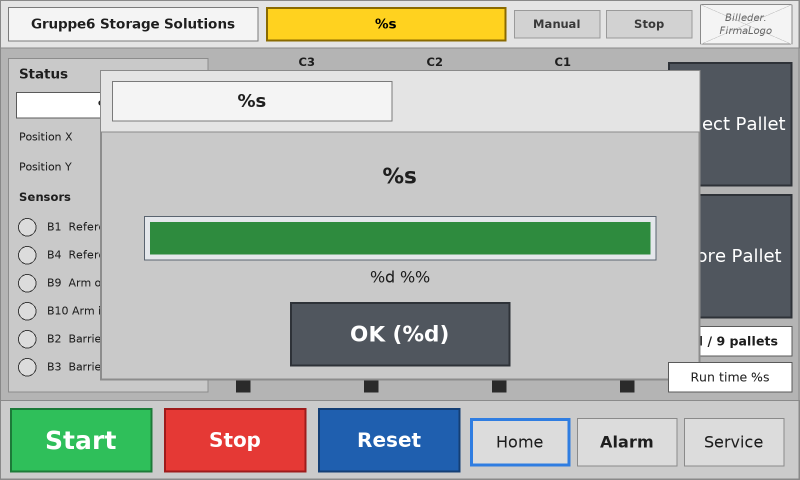
VISUALIZATION Start  // 800x480
    Rectangle (0,0 800x480)
    Rectangle (0,0 800x48)
    Rectangle (8,7 250x34), "Gruppe6 Storage Solutions"
    Rectangle (266,7 150x34), "OP031 Warehouse"
    Rectangle (514,10 86x28), "Manual", colour toggle: MAIN.isManualMode
    Rectangle (606,10 86x28), "Stop", colour toggle: MAIN.isStop
    Rectangle (0,400 800x80)
    RoundedRectangle (10,408 142x64), "Start"
        OnMouseUp: execute { MAIN.isStop := FALSE; }
    RoundedRectangle (164,408 142x64), "Stop"
        OnMouseUp: execute { MAIN.isStop := TRUE; }
    RoundedRectangle (318,408 142x64), "Reset"
        OnMouseUp: execute {
            MAIN.resetRequest := TRUE;   // everything back to Step_10, then homing
        }
    Rectangle (470,418 100x48), "Home"
        OnMouseUp: change screen: Start
    Rectangle (684,418 100x48), "Service"
        OnMouseUp: change screen: Service
    Rectangle (8,58 200x334)
    Rectangle (16,62 184x24), "Status"
    Rectangle (16,124 84x26), "Position X"
    Rectangle (100,124 100x26), "%d", text variable: MAIN.currentPosX
    Rectangle (16,154 84x26), "Position Y"
    Rectangle (100,154 100x26), "%d", text variable: MAIN.currentPosY
    Rectangle (16,186 184x22), "Sensors"
    Ellipse (18,218 18x18), colour toggle: MAIN.B1
    Rectangle (44,214 160x26), "B1 Reference X"
    Ellipse (18,246 18x18), colour toggle: MAIN.B4
    Rectangle (44,242 160x26), "B4 Reference Y (top)"
    Ellipse (18,274 18x18), colour toggle: MAIN.B9
    Rectangle (44,270 160x26), "B9 Arm out"
    Ellipse (18,302 18x18), colour toggle: MAIN.B10
    Rectangle (44,298 160x26), "B10 Arm in"
    Ellipse (18,330 18x18), colour toggle: MAIN.B2
    Rectangle (44,326 160x26), "B2 Barrier in (free)"
    Ellipse (18,358 18x18), colour toggle: MAIN.B3
    Rectangle (44,354 160x26), "B3 Barrier out (free)"
    Rectangle (236,74 14x318)
    Rectangle (364,74 14x318)
    Rectangle (492,74 14x318)
    Rectangle (620,74 14x318)
    Rectangle (236,150 398x10)
    Rectangle (640,120 24x24), "R3"
    Rectangle (236,250 398x10)
    Rectangle (640,220 24x24), "R2"
    Rectangle (236,350 398x10)
    Rectangle (640,320 24x24), "R1"
    Rectangle (277,52 60x20), "C3"
    Rectangle (405,52 60x20), "C2"
    Rectangle (533,52 60x20), "C1"
    Rectangle (265,110 84x40), colour toggle: MAIN.slotOccupied[3,3]
    Rectangle (272,101 70x9), colour toggle: MAIN.slotOccupied[3,3]
    Rectangle (393,110 84x40), colour toggle: MAIN.slotOccupied[2,3]
    Rectangle (400,101 70x9), colour toggle: MAIN.slotOccupied[2,3]
    Rectangle (521,110 84x40), colour toggle: MAIN.slotOccupied[1,3]
    Rectangle (528,101 70x9), colour toggle: MAIN.slotOccupied[1,3]
    Rectangle (265,210 84x40), colour toggle: MAIN.slotOccupied[3,2]
    Rectangle (272,201 70x9), colour toggle: MAIN.slotOccupied[3,2]
    Rectangle (393,210 84x40), colour toggle: MAIN.slotOccupied[2,2]
    Rectangle (400,201 70x9), colour toggle: MAIN.slotOccupied[2,2]
    Rectangle (521,210 84x40), colour toggle: MAIN.slotOccupied[1,2]
    Rectangle (528,201 70x9), colour toggle: MAIN.slotOccupied[1,2]
    Rectangle (265,310 84x40), colour toggle: MAIN.slotOccupied[3,1]
    Rectangle (272,301 70x9), colour toggle: MAIN.slotOccupied[3,1]
    Rectangle (393,310 84x40), colour toggle: MAIN.slotOccupied[2,1]
    Rectangle (400,301 70x9), colour toggle: MAIN.slotOccupied[2,1]
    Rectangle (521,310 84x40), colour toggle: MAIN.slotOccupied[1,1]
    Rectangle (528,301 70x9), colour toggle: MAIN.slotOccupied[1,1]
    RoundedRectangle (668,62 124x124), "Select Pallet"
        OnMouseUp: execute {
            MAIN.awaitingUserInput := TRUE;   // tell the SFC (Step_10): the operator wants to retrieve a pallet
        }
        OnMouseUp: OpenDialog Dialog=SelectPalletDialog, OpenModal=True, OpenCentered=True
    RoundedRectangle (668,194 124x124), "Store Pallet", colour toggle: MAIN.isStorageFull
        OnMouseUp: execute {
            MAIN.storeRequest := TRUE;   // run the pallet in on the conveyor (to B2) and store it in the rack
        }
    Image (700,4 92x40), image: Billeder.FirmaLogo
    Rectangle (16,92 184x26), "%s", text variable: MAIN.statusText
    Rectangle (668,326 124x30), "%d / 9 pallets", text variable: MAIN.palletCount
    Rectangle (100,70 600x310), invisible if: MAIN.hideStorageFull, input disabled if: MAIN.hideStorageFull
    Rectangle (100,70 600x62), invisible if: MAIN.hideStorageFull, input disabled if: MAIN.hideStorageFull
    Rectangle (112,81 200x40), "Warning", invisible if: MAIN.hideStorageFull, input disabled if: MAIN.hideStorageFull
    Rectangle (528,84 160x34), "Storage full", invisible if: MAIN.hideStorageFull, input disabled if: MAIN.hideStorageFull
    Rectangle (120,180 560x60), "Storage is full, remove pallets first", invisible if: MAIN.hideStorageFull, input disabled if: MAIN.hideStorageFull
    RoundedRectangle (290,288 220x64), "OK", invisible if: MAIN.hideStorageFull, input disabled if: MAIN.hideStorageFull
        OnMouseUp: execute {
            MAIN.showStorageFull := FALSE;   // close the message
        }
    Rectangle (100,70 600x310), invisible if: MAIN.hideProgress, input disabled if: MAIN.hideProgress
    Rectangle (100,70 600x62), invisible if: MAIN.hideProgress, input disabled if: MAIN.hideProgress
    Rectangle (112,81 280x40), "%s", text variable: MAIN.progressTitle, invisible if: MAIN.hideProgress, input disabled if: MAIN.hideProgress
    Rectangle (120,148 560x56), "%s", text variable: MAIN.progressText, invisible if: MAIN.hideProgress, input disabled if: MAIN.hideProgress
    Rectangle (144,216 512x44), invisible if: MAIN.hideProgress, input disabled if: MAIN.hideProgress
    Rectangle (150,222 25x32), invisible if: MAIN.progressHide[1], input disabled if: MAIN.progressHide[1]
    Rectangle (175,222 25x32), invisible if: MAIN.progressHide[2], input disabled if: MAIN.progressHide[2]
    Rectangle (200,222 25x32), invisible if: MAIN.progressHide[3], input disabled if: MAIN.progressHide[3]
    Rectangle (225,222 25x32), invisible if: MAIN.progressHide[4], input disabled if: MAIN.progressHide[4]
    Rectangle (250,222 25x32), invisible if: MAIN.progressHide[5], input disabled if: MAIN.progressHide[5]
    Rectangle (275,222 25x32), invisible if: MAIN.progressHide[6], input disabled if: MAIN.progressHide[6]
    Rectangle (300,222 25x32), invisible if: MAIN.progressHide[7], input disabled if: MAIN.progressHide[7]
    Rectangle (325,222 25x32), invisible if: MAIN.progressHide[8], input disabled if: MAIN.progressHide[8]
    Rectangle (350,222 25x32), invisible if: MAIN.progressHide[9], input disabled if: MAIN.progressHide[9]
    Rectangle (375,222 25x32), invisible if: MAIN.progressHide[10], input disabled if: MAIN.progressHide[10]
    Rectangle (400,222 25x32), invisible if: MAIN.progressHide[11], input disabled if: MAIN.progressHide[11]
    Rectangle (425,222 25x32), invisible if: MAIN.progressHide[12], input disabled if: MAIN.progressHide[12]
    Rectangle (450,222 25x32), invisible if: MAIN.progressHide[13], input disabled if: MAIN.progressHide[13]
    Rectangle (475,222 25x32), invisible if: MAIN.progressHide[14], input disabled if: MAIN.progressHide[14]
    Rectangle (500,222 25x32), invisible if: MAIN.progressHide[15], input disabled if: MAIN.progressHide[15]
    Rectangle (525,222 25x32), invisible if: MAIN.progressHide[16], input disabled if: MAIN.progressHide[16]
    Rectangle (550,222 25x32), invisible if: MAIN.progressHide[17], input disabled if: MAIN.progressHide[17]
    Rectangle (575,222 25x32), invisible if: MAIN.progressHide[18], input disabled if: MAIN.progressHide[18]
    Rectangle (600,222 25x32), invisible if: MAIN.progressHide[19], input disabled if: MAIN.progressHide[19]
    Rectangle (625,222 25x32), invisible if: MAIN.progressHide[20], input disabled if: MAIN.progressHide[20]
    Rectangle (144,264 512x26), "%d %%", text variable: MAIN.progressPercent, invisible if: MAIN.hideProgress, input disabled if: MAIN.hideProgress
    RoundedRectangle (290,302 220x64), "OK (%d)", text variable: MAIN.okCountdown, invisible if: MAIN.hideProgressOk, input disabled if: MAIN.hideProgressOk
        OnMouseUp: execute {
            MAIN.retrievePhase := 0; MAIN.storePhase := 0;   // close the progress box
        }
    Rectangle (577,418 100x48), "Alarm", colour toggle: MAIN.isAlarm
        OnMouseUp: change screen: Alarm
    Rectangle (668,362 124x30), "Run time %s", text variable: MAIN.runTimeText
    Rectangle (266,7 240x34), "%s", text variable: MAIN.alarmBannerText, invisible if: MAIN.hideAlarmBanner, input disabled if: MAIN.hideAlarmBanner
        OnMouseUp: change screen: Alarm
END_VISUALIZATION

(* stored: Version 1.1.0.1, ProductVersion 3.1.4024.12
   Visu Start: Id {1ddcc670-8b4f-4c7f-936e-57019fb79669} *)
